PROGRAM main
  VAR
    S1 AT %IX0.0 : BOOL; (* barrera de entrada: entra un auto *)
    S2 AT %IX0.1 : BOOL; (* barrera de salida: sale un auto *)
    H1 AT %QX0.0 : BOOL; (* verde: hay lugar *)
    H2 AT %QX0.1 : BOOL; (* amarillo: lleno *)
    F_ENTRA      : R_TRIG;
    F_SALE       : R_TRIG;
    AUTOS        : INT; (* autos adentro *)
    LIBRES       : INT; (* lugares libres *)
    ENTRA        : BOOL; (* flanco de S1 *)
    SALE         : BOOL; (* flanco de S2 *)
    HAY_LUGAR    : BOOL; (* AUTOS < capacidad *)
    HAY_AUTOS    : BOOL; (* AUTOS > 0 *)
  END_VAR
  VAR  (* added by the conversion: wires and edge detectors of the diagram *)
    _ADD10_OUT : INT;
    _SEL7_OUT : INT;
    _SUB17_OUT : INT;
    _SEL14_OUT : INT;
    _SUB21_OUT : INT;
    _GT25_OUT : BOOL;
    _LE29_OUT : BOOL;
  END_VAR

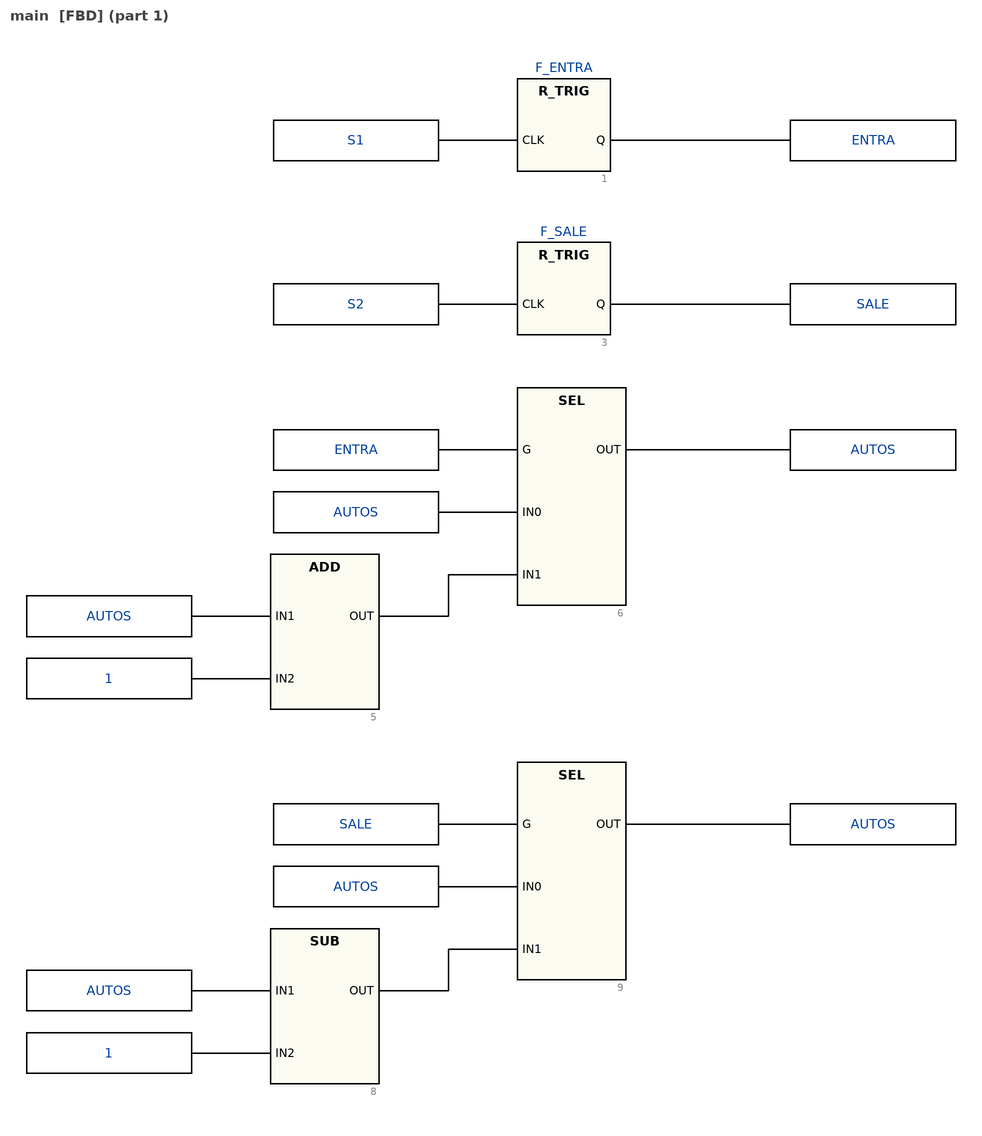
(* FBD diagram, written out as Structured Text *)
F_ENTRA(CLK := S1);
ENTRA := F_ENTRA.Q;
F_SALE(CLK := S2);
SALE := F_SALE.Q;
_ADD10_OUT := AUTOS + 1;
_SEL7_OUT := SEL(ENTRA, AUTOS, _ADD10_OUT);
AUTOS := _SEL7_OUT;
_SUB17_OUT := AUTOS - 1;
_SEL14_OUT := SEL(SALE, AUTOS, _SUB17_OUT);
AUTOS := _SEL14_OUT;
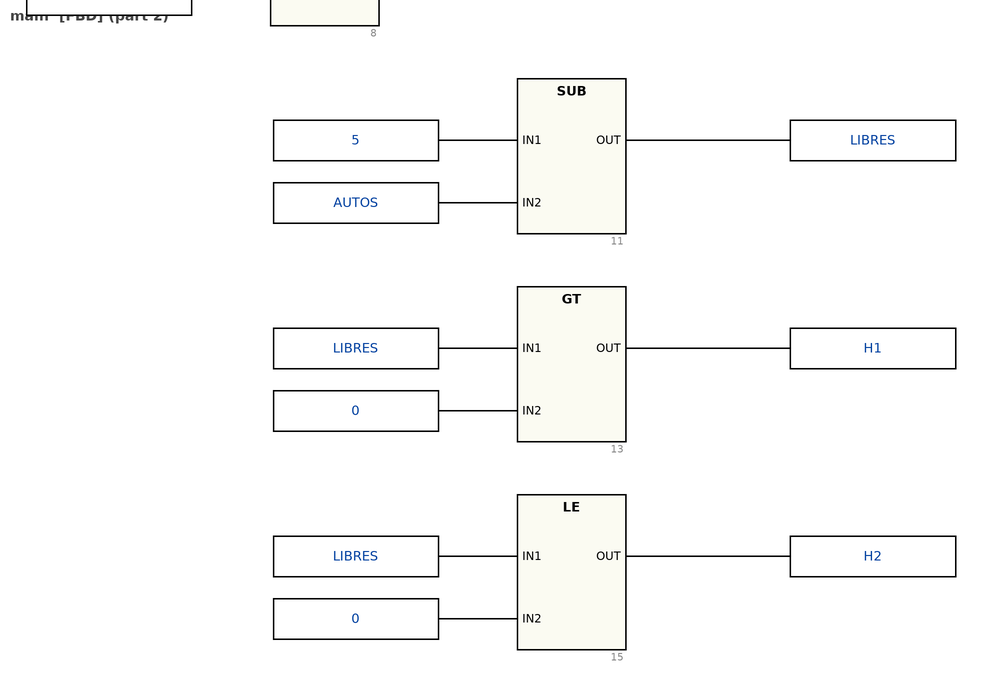
_SUB21_OUT := 5 - AUTOS;
LIBRES := _SUB21_OUT;
_GT25_OUT := LIBRES > 0;
H1 := _GT25_OUT;
_LE29_OUT := LIBRES <= 0;
H2 := _LE29_OUT;
END_PROGRAM
